// Sortie numérique, type 2 (docs/03 § 3.2)
FUNCTION_BLOCK FB_DigitalOutput EXTENDS FB_ObjectBase
VAR
    _bCmd : BOOL;
    _fPulseMs : LREAL;
    _fElapsed : LREAL;
END_VAR

METHOD PROTECTED _OnConfigure : BOOL
_OnConfigure := F_SignalValid(_refCfg.aSignal[1], E_SignalKind.DO);
END_METHOD

METHOD PROTECTED _DefaultTimeoutMs : UDINT
VAR_INPUT
    nAction : UINT;
END_VAR
IF nAction = GVL_Catalog.DigitalOutput_Impulsion THEN
    _DefaultTimeoutMs := LREAL_TO_UDINT(_ParamReal(1, _refCfg.aParam[2])) + 1000;
ELSE
    _DefaultTimeoutMs := 0;
END_IF
END_METHOD

METHOD PROTECTED _ValidateParams : BOOL
VAR_INPUT
    nAction : UINT;
END_VAR
_ValidateParams := nAction <> GVL_Catalog.DigitalOutput_Impulsion OR _ParamReal(1, _refCfg.aParam[2]) >= 1.0;
END_METHOD

METHOD PROTECTED _OnStart : E_ActStatus
VAR_INPUT
    nAction : UINT;
END_VAR
CASE nAction OF
    GVL_Catalog.DigitalOutput_Activer:
        _bCmd := TRUE;
        _OnStart := E_ActStatus.Done;
    GVL_Catalog.DigitalOutput_Desactiver:
        _bCmd := FALSE;
        _OnStart := E_ActStatus.Done;
    GVL_Catalog.DigitalOutput_Impulsion:
        _fPulseMs := LIMIT(1.0, _ParamReal(1, _refCfg.aParam[2]), 60000.0);
        _fElapsed := 0;
        _bCmd := TRUE;
        _OnStart := E_ActStatus.Busy;
ELSE
    _OnStart := E_ActStatus.Error;
END_CASE
END_METHOD

METHOD PROTECTED _OnCycle : E_ActStatus
VAR_INPUT
    nAction : UINT;
END_VAR
_fElapsed := _fElapsed + F_CycleMs();
IF _fElapsed >= _fPulseMs THEN
    _bCmd := FALSE;
    _OnCycle := E_ActStatus.Done;
ELSE
    _OnCycle := E_ActStatus.Busy;
END_IF
END_METHOD

METHOD PROTECTED _SafeState
CASE LREAL_TO_INT(_refCfg.aParam[3]) OF
    0: _bCmd := FALSE;
    1: _bCmd := TRUE;
END_CASE                            // 2 : maintien
END_METHOD

METHOD PROTECTED _WriteHw
F_WriteDO(_refCfg.aSignal[1], _bCmd XOR (_refCfg.aParam[1] = 1));
END_METHOD

METHOD PROTECTED _Publish
_stStatus.aValue[1] := BOOL_TO_LREAL(_bCmd);
END_METHOD

END_FUNCTION_BLOCK

(* stored: Version 1.1.0.1, ProductVersion 3.1.4024.12
   POU FB_DigitalOutput: Id {70e1d49b-9dcb-57f8-9796-be045f1bf688}, SpecialFunc None
   Method _OnConfigure: Id {78f26ede-9171-5b1b-8255-2ecb3758e185}
   Method _DefaultTimeoutMs: Id {f98d6076-6952-5ef1-b7d0-54a0a26f9815}
   Method _ValidateParams: Id {dc67c4ce-47c5-5f75-b235-14fe1ef5952c}
   Method _OnStart: Id {2ffa91fa-1fae-5520-a4fc-ff4939ba8ebb}
   Method _OnCycle: Id {7ffd0e05-afbf-5c8a-8b04-0fa6f0c43e18}
   Method _SafeState: Id {a2f5e23c-49a2-53d7-b837-0958787c7729}
   Method _WriteHw: Id {4fe98c43-f91c-578c-990f-0786fe27a1cd}
   Method _Publish: Id {c7db503d-cdcf-5946-a05e-bfa5e495e9b8} *)
